(* IEC 61131-3 sources: CS_4_Aufzugsteuerung/src/Stations/CP112/Steuerung/Class/SdiasSafetyManagerFSoE (part 2) *)

            LastRequest := _WriteSysTime;

            //copy SDO into write-buffer
            ToStdLib.MemCpy(dest := #p_Handle_SDO_Write^.SDOStructure, source := #StandardRequest, size := (sizeof(SDOHeader.StdHeader.CRC) + StandardRequest.SDOHeader.Len));

            //mark SDO data as valid
            p_Handle_SDO_Write^.us_Status := SAFETY_SDO_DATA_VALID;

            if ( pISafety^.udVersion >= 16#1001 ) then
              SAFETY_iPushSafetyTask();
            end_if;

            SDOTimeMark       := ops.tAbsolute;
            ud_LastSetSysTime := ops.tAbsolute;
            eResponseState    := _wait;

            // check timeout
          elsif ((ops.tAbsolute - SDOTimeMark) > SDIAS_SAFTEY_SDO_RESPONSE_TIMEOUT) & (eResponseState <> _valid) then
            LogError("@029F (SdiasSafetyManagerFSoE::InitModule) Timeout while waiting for the SDO Send buffer to get ready (set system time)");
            eInitSSWErrorStep := eInitSSW;
            eInitSSW          := _InitError;
          end_if;

      //*****************************************************
        _wait: // wait for response

          //check id sdo sending was ok
          if ( p_Handle_SDO_Read^.us_Status = SAFETY_SDO_DATA_VALID ) then

            //calculate length of SDO
            us_SDO_length := sizeof(SDOHeader.StdHeader.CRC) + p_Handle_SDO_Read^.SDOStructure.SDOHeader.StdHeader.Len;

            //copy SDO without first byte (=status byte)
            ToStdLib.MemCpy(dest := p_SDOOutputBuffer, source := #p_Handle_SDO_Read^.SDOStructure, size := us_SDO_length );

            //mark data as received
            p_Handle_SDO_Read^.us_Status := SAFETY_SDO_NO_DATA;

            //check, if it's our answer
            if ((p_SDOOutputBuffer^.SDOHeader.StdHeader.Typ$USINT AND SBF_SSDO_MASK_TYPE)$t_SafetyFrameType = SDO_STD) then
              StandardResponse := (p_SDOOutputBuffer$^StandardFrameType)^;
              if StandardResponse.SDOHeader.SeqNr = (StandardSeqNr OR 16#80) then
                if LastRequest = _WriteSysTime then
                  // delete request
                  LastRequest           := _NoOpenRequest;
                  ud_AsyComRetryCounter := 0; // reset retry counter
                  eResponseState        := _valid;
                  // if returnvalue is 34 (E_SM_SSDO_INVALID_VIRTADDR) the virtual address is not supported by firmware
                  if StandardResponse.aData[0] <> 34 then
                    //virtual adress for write of timestamp is supported
                    b_SetSysTime := TRUE;
                  else
                    b_SetSysTime := FALSE;
                  end_if;
                else
                  LogError("@025A (SdiasSafetyManagerFSoE::InitModule) SDO Receive: Invalid standard frame response.");
                  eInitSSWErrorStep := eInitSSW;
                  eInitSSW          := _InitError;
                end_if;

                // if request is deleted, increase sequence number to set next request
                if LastRequest = _NoOpenRequest then
                  if StandardSeqNr < 16#7F then
                    StandardSeqNr += 1;
                  else
                    StandardSeqNr := 0;
                  end_if;
                end_if;
              else
                LogError("@025B (SdiasSafetyManagerFSoE::InitModule) SDO Receive: Invalid sequence number in Standard SDO response.");
                LogValue("expected: 0x{0} / received: 0x{1}", Value:=(StandardSeqNr OR 16#80), Value2:=StandardResponse.SDOHeader.SeqNr);
                eInitSSWErrorStep := eInitSSW;
                eInitSSW          := _InitError;
              end_if;
            else
              // ignore non-standard frames => the module may try to distribute it's configuration
            end_if;
          end_if;

          // check timeout
          if ((ops.tAbsolute - SDOTimeMark) > SDIAS_SAFTEY_SDO_RESPONSE_TIMEOUT) & (eResponseState <> _valid) then
            LogError("@02A1 (SdiasSafetyManagerFSoE::InitModule) SDO Response timeout while waiting for the module configuration.");
            eInitSSWErrorStep := eInitSSW;
            eInitSSW          := _InitError;
          end_if;
      //*****************************************************
        _valid:
          eInitSSW        := _DisablePLL;
          eResponseState  := _idle;
      //*****************************************************
      end_case;

//**********************************************************************************************************************************************************
    _DisablePLL: // disable the PLL
      TmpRetCode := BusConfigWrite(Offset:=SDIAS_SAFETY_PLL_OFFSET + t_PllRegister.StatusControl, Length:=sizeof(sPllRegister.StatusControl), pData:=#sPllRegister.StatusControl, IsControlAccess:=TRUE);

      if TmpRetCode = READY then
        eInitSSW := _GetPLLSettings;
      elsif TmpRetCode = ERROR then
        eInitSSW := _InitError;
      end_if;

//**********************************************************************************************************************************************************
    _GetPLLSettings: // get the actual PLL settings
      TmpRetCode := BusConfigRead(Offset:=SDIAS_SAFETY_PLL_OFFSET, Length:=sizeof(sPllRegister), pData:=#sPllRegister, IsControlAccess:=TRUE);

      if TmpRetCode = READY then
        // get bus cycle time for the PLL settings
        MyPara.uiCmd     := _BUS_IF_GET_BUSCYCLE_TIME;

        ToBusInterface.NewInst(pPara:=#MyPara, pResult:=#MyResult);
        if MyResult.aData[0]$t_GetBusCycleTime.retcode = _BUS_IF_RETVAL_OK then
          udBusTime       := MyResult.aData[0]$t_GetBusCycleTime.udBusCycleTime;
        else
          // use this just to have
          udBusTime := 1000;
          LogError("@02AA (SdiasSafetyManagerFSOE::InitModule) Failed to get bus cycle settings BusInterface.");
        end_if;

        udBusTime_us := udBusTime / 1000;

        // settings for pll
        sPllRegister.SystemPeriodTime           := udBusTime / 10;            // convert to 10*ns
        sPllRegister.StatusControl              := 0;
        sPllRegister.StatusControl.SyncEnable   := 1;
        sPllRegister.PeriodDivider              := to_usint(udBusTime_us / 1000);  // Bustime / 1ms to get divider (0 and 1 gets the same result)
        //sPllRegister.CompensationDelay // Keep value
        sPllRegister.SyncOut0.Offset            := 0;
        sPllRegister.SyncOut0.PeriodMultiplier  := to_usint(1000 / udBusTime_us);  // 1ms / Bustime to get multiplier (0 and 1 gets the same result);
        sPllRegister.SyncOut0.SyncStartDelay    := 0;
        sPllRegister.SyncOut0.ControlStatusRegister.SyncOutEnable     := 1;
        sPllRegister.SyncOut0.ControlStatusRegister.StartDelayEnable  := 0;
        if sPllRegister.PeriodDivider <= 1 then
          // no divider use system sync
          sPllRegister.SyncOut0.ControlStatusRegister.SyncSelector       := 1;  // no divider use system sync
        else
          // a divider is defined -> use it
          sPllRegister.SyncOut0.ControlStatusRegister.SyncSelector       := 0;
        end_if;

        eInitSSW := _ConfigurePLL;
      elsif TmpRetCode = ERROR then
        eInitSSW := _InitError;
      end_if;

//**********************************************************************************************************************************************************
    _ConfigurePLL:
      TmpRetCode := BusConfigWrite(Offset:=SDIAS_SAFETY_PLL_OFFSET, Length:=sizeof(sPllRegister), pData:=#sPllRegister, IsControlAccess:=TRUE);

      if TmpRetCode = READY then

        eInitSSW := _ConfigureTripleBufferAnalogReadData;
      elsif TmpRetCode = ERROR then
        eInitSSW := _InitError;
      end_if;

//**********************************************************************************************************************************************************
    _ConfigureTripleBufferAnalogReadData:

      //check if config from triple buffer for analog data is necessary
      if usAnalogInputByteSize then

        // configure the triple buffer - the required bytes are passed to the FPGA.
        sAnalogTripleBufferConfig.usSizeuCtoCPU := usAnalogInputByteSize - sizeof(USINT); //-1 byte for messagecounter
        sAnalogTripleBufferConfig.usSizeCPUtouC := 0; //Analog write when supported

        TmpRetCode := BusConfigWrite(Offset:=SBF_OFFSET_ANALOG_VALUE_TRIPLE_PUFFER_SWITCH_OFFSET_WR_1, Length:=sizeof(sAnalogTripleBufferConfig), pData:=#sAnalogTripleBufferConfig, IsControlAccess:=FALSE);

        if TmpRetCode = READY then
          eInitSSW := _ConfigureFastTripleBuffer;
        elsif TmpRetCode = ERROR then
          eInitSSW := _InitError;
        end_if;
      else
        eInitSSW := _ConfigureFastTripleBuffer;
      end_if;

//**********************************************************************************************************************************************************
    _ConfigureFastTripleBuffer:

      //check if init from triple buffer is necessary
      if uiPDOReadSizeFastUnsafeVar <> 0 |
        uiPDOWriteSizeFastUnsafeVar <> 0 then

        // configure the triple buffer - the required bytes are passed to the FPGA.
        sFastTripleBufferConfig.SizeuCtoCPU := uiPDOReadSizeFastUnsafeVar$USINT - 1;
        sFastTripleBufferConfig.SizeCPUtouC := uiPDOWriteSizeFastUnsafeVar$USINT - 1;

        TmpRetCode := BusConfigWrite(Offset:=SBF_OFFSET_FAST_UNSAFE_BUFFER_CONFIG, Length:=sizeof(sFastTripleBufferConfig), pData:=#sFastTripleBufferConfig, IsControlAccess:=FALSE);

        if TmpRetCode = READY then
          eInitSSW := _Finished;
        elsif TmpRetCode = ERROR then
          eInitSSW := _InitError;
        end_if;
      else
        eInitSSW := _Finished;
      end_if;

//**********************************************************************************************************************************************************
    _Finished:
      //Only set online here to 1 if we don't have to adjust the the triple buffer config, otherwise online will be set in cyclic after correcting the triple buffer config
      if b_ModuleAccessReady & (bWriteAnalogTripleBufferConfig = FALSE) then
        Online := 1;
      end_if;

      eInitSSW          := _PrepareInit;
      ModuleInitState   := READY;

#ifdef SAFETY_iDisableNonClassCommunication
      if ( pISafety^.udVersion >= 16#1002 ) then
        SAFETY_iDisableNonClassCommunication(uiMaster:=0, pucNode:=p_ObjectPath, uiDisable:=0);
      end_if;
#endif

//**********************************************************************************************************************************************************
    _InitError:
      eInitSSW          := _PrepareInit;
      ModuleInitState   := ERROR;

#ifdef SAFETY_iDisableNonClassCommunication
      if ( pISafety^.udVersion >= 16#1002 ) then
        SAFETY_iDisableNonClassCommunication(uiMaster:=0, pucNode:=p_ObjectPath, uiDisable:=0);
      end_if;
#endif

//**********************************************************************************************************************************************************
  end_case;

END_FUNCTION

FUNCTION VIRTUAL GLOBAL SdiasSafetyManagerFSoE::ClassSvr::NewInst
  VAR_INPUT
    pPara 	: ^CmdStruct;
    pResult 	: ^results;
  END_VAR
  VAR_OUTPUT
    ret_code 	: iprStates;
  END_VAR
  VAR
    i                 : UDINT;
    pSafetyModuleInfo : ^t_SdiasSafetyModuleInfo;
    MyPara 	          : CmdStruct;
    MyResult          : Results;
    HBGPlace          : UDINT;
    bRequiredError    : BOOL;
    bHWConfigError    : BOOL;

    pStr_HWTRequested     : ^CHAR;
    tmpplace      : USINT;
    pStr_HWTreeEntry : ^CHAR;
    usNextPlace   : USINT;
    pNewElement   : t_pHWCGetHardwareDiagnosisOutDynExt;
    usTmpAnalogInputByteSize : USINT;
  END_VAR

  ret_code := ERROR;

  CASE pPara^.uiCmd OF

//*****************************************************************************
//**  COMMANDS FROM BUS INTERFACE                                            **
//*****************************************************************************

//**********************************************************************************************************************************************************
    _BUS_IF_INIT_ACCESSES:
      // is called until the module is ready or in error state (only done once when no accesses have been created yet)
      ret_code := InitAccess();

//**********************************************************************************************************************************************************
    _BUS_IF_INIT_MODULE:
      // is called until the module is ready or in error state (done every time the module is connected)
      ret_code := InitModule();

//**********************************************************************************************************************************************************
    _BUS_IF_SDO_RESPONSE:
      // check if the command matches the one we're waiting for
      if (pPara^.aPara[0] = LastSDO.Command) &
         (pPara^.aPara[1] = LastSDO.Offset)  &
         (pPara^.aPara[2] = LastSDO.Length) then

        if pPara^.aPara[3]$iprStates = READY then
          if (LastSDO.Command = _BUS_IF_READ_VIA_SDO) then
            if (LastSDO.Offset = SBF_OFFSET_IO_MODULE_IDS) then
              if eResponseState = _wait then
                if pPara^.aPara[5] = LastSDO.Length then
                  if pPara^.aPara[4] then
                    // all parameters are fine, so we're ready
                    ret_code := READY;

                    _memcpy(ptr1:=#aModuleIDs, ptr2:=pPara^.aPara[4]$pVoid, cntr:=LastSDO.Length);

                    bRequiredError := FALSE;
                    bHWConfigError := FALSE;

                    //Set byte size of analog inputs to zero (will be summarized with every analog module)
                    usTmpAnalogInputByteSize := 0;

                    // search for a HBG in the module IDs
                    HBGPlace := SDIAS_SAFETY_INVALID_MAX_PLACE;
                    for i := 0 to 16 do
                      if (aModuleIDs[i] AND SDIAS_SAFETY_MODULE_ID_BUS_MASK) = SDIAS_SAFETY_MODULE_ID_CAN_BUS_MASK then
                        HBGPlace := i;
                        exit;
                      end_if;
                    end_for;

                    // now we got the module IDs according to the safety cpu => check if it matches our configuration (only available on newer firmware versions)
                    if b_GotOptionalSettings then
                      pSafetyModuleInfo := #aSafetyModuleInfo[0];

                      // always the same command
                      MyPara.uiCmd := SDIAS_SET_CLASS_STATE;

                      for i := 0 to 15 do
                        MyPara.aPara[1] := aModuleIDs[i];

                        // if a required module is not matching => required error
                        if pSafetyModuleInfo^.sdRequired & (aModuleIDs[i] <> pSafetyModuleInfo^.usExpectedDeviceID) then
                          MyPara.aPara[0] := _RequiredError$DINT;
                          bRequiredError := TRUE;
                          if aModuleIDs[i] = SDIAS_SAFETY_INVALID_DEVICE_ID then
                            LogValue("@02AB (SdiasSafetyManagerFSoE::ClassSvr::NewInst) No safety IO module at required place {0}", Value:=i);
                          else
                            LogValue("@02AC (SdiasSafetyManagerFSoE::ClassSvr::NewInst) Wrong safety IO module at required place {0}", Value:=i);
                          end_if;

                        // check if the configuration in the safety designer matches the configuration in the hardware classes
                        elsif pSafetyModuleInfo^.usExpectedDeviceID = OptionalSettings.ModuleIDsConfigured[i] then
                          // if it's an invalid device ID, it's only allowed if there is no module
                          if pSafetyModuleInfo^.usExpectedDeviceID = SDIAS_SAFETY_INVALID_DEVICE_ID then
                            if aModuleIDs[i] = SDIAS_SAFETY_INVALID_DEVICE_ID then
                              // correct (no module configured and no module found)
                              MyPara.aPara[0] := _ClassOk$DINT;  // this value is not being written to the module since if the ID is 0, there is also no this pointer to call the newinst
                            elsif (i <> HBGPlace) then
                              // no module configured but a module has been found at this place
                              LogValue("@02AD (SdiasSafetyManagerFSoE::ClassSvr::NewInst) No module configured in hardware classes and safety designer but found module at place {0}", Value:=i);
                              MyPara.aPara[0] := _WrongHardware$DINT; // again no object to write this value to
                              bHWConfigError := TRUE;
                            end_if;

                          // now check if we got the expected ID at this position
                          elsif aModuleIDs[i] = pSafetyModuleInfo^.usExpectedDeviceID then
                            // correct module
                            MyPara.aPara[0] := _ClassOk$DINT;

                            //Check if this is an analog module
                            if pSafetyModuleInfo^.usAnalogInputByteSize then
                              //Increase our byte size --> mabye we need to refresh the byte size in the tripple buffer of the analog values if the amount of configured modules
                              //differs to the amount of available modules on the hardware (e.g optional modules)
                              if usTmpAnalogInputByteSize = 0 then
                                usTmpAnalogInputByteSize += pSafetyModuleInfo^.usAnalogInputByteSize + sizeof(USINT);  //Add one byte for message counter if not added yet (first byte of analog input buffer is messagecounter)
                              else
                                usTmpAnalogInputByteSize += pSafetyModuleInfo^.usAnalogInputByteSize;
                              end_if;
                            end_if;

                            // if this module is optional
                          elsif OptionalSettings.OptionalFlagsIOModules AND (1 SHL i) then
                            // if it's a blank module
                            if aModuleIDs[i] = SDIAS_SAFETY_MODULE_ID_BLANK_MODULE then
                              // ok: blank is allowed at optional place
                              MyPara.aPara[0] := _NoHardware$DINT;

                              // don't send the blank-module ID
                              MyPara.aPara[1] := SDIAS_SAFETY_INVALID_DEVICE_ID;
                            else
                              if aModuleIDs[i] = SDIAS_SAFETY_INVALID_DEVICE_ID then
                                // ok: no module instead of the configured one (allowed since it's the last module. no more modules possible after an invalid device id)
                                MyPara.aPara[0] := _NoHardware$DINT;

                              //optional module, maybe this module is the HBG itself
                              elsif (HBGPlace <> SDIAS_SAFETY_INVALID_MAX_PLACE) & (i = HBGPlace) then

                                //OK: optional module is not available and this one is the HBG
                                MyPara.aPara[0] := _NoHardware$DINT;
                                MyPara.aPara[1] := SDIAS_SAFETY_INVALID_DEVICE_ID;
                              else
                                // wrong module detected
                                MyPara.aPara[0] := _WrongHardware$DINT;
                                bHWConfigError := TRUE;
                                LogValue("@02AE (SdiasSafetyManagerFSoE::ClassSvr::NewInst) Wrong safety IO module at place {0}. (configured as optional)", Value:=i);
                              end_if;
                            end_if;
                          else
                            // the module id does not match (missing or wrong module)
                            if aModuleIDs[i] = SDIAS_SAFETY_INVALID_DEVICE_ID then
                              MyPara.aPara[0] := _NoHardware$DINT;
                            else
                              MyPara.aPara[0] := _WrongHardware$DINT;
                            end_if;

                            // check if it's required
                            if MyPara.aPara[0] = _NoHardware$DINT then
                              LogValue("@02AF (SdiasSafetyManagerFSoE::ClassSvr::NewInst) No safety IO module at place {0}.", Value:=i);
                            else
                              LogValue("@02B0 (SdiasSafetyManagerFSoE::ClassSvr::NewInst) Wrong safety IO module at place {0}.", Value:=i);
                            end_if;

                            bHWConfigError := TRUE;
                          end_if;
                        else
                          // the configuration in the safety designer differs from the configuration via the hardware classes

                          // if the available hardware matches the safety designer configuration and there is no module (only in hw class configuration)
                          if (OptionalSettings.ModuleIDsConfigured[i] = SDIAS_SAFETY_INVALID_DEVICE_ID) &
                             ((aModuleIDs[i] = SDIAS_SAFETY_INVALID_DEVICE_ID) | (i = HBGPlace)) &
                             (pSafetyModuleInfo^.usExpectedDeviceID <> SDIAS_SAFETY_INVALID_DEVICE_ID) then
                            // that's allowed
                            LogValue("@02B1 (SdiasSafetyManagerFSoE::ClassSvr::NewInst) Module in hardware class configuration which is neither available physically nor in safety designer configuration at place {0}", Value:=i);
                            MyPara.aPara[0] := _NoHardware$DINT;

                          else
                            // in all other cases, it isn't
                            LogValue("@02B2 (SdiasSafetyManagerFSoE::ClassSvr::NewInst) Module in hardware class configuration differs from safety designer configuration at place {0}", Value:=i);
                            MyPara.aPara[0] := _InvalidConfguration$DINT;
                            bHWConfigError := TRUE;
                          end_if;
                        end_if;

                        if pSafetyModuleInfo^.pThis then
                          pSafetyModuleInfo^.pThis^.NewInst(#MyPara, #MyResult);
                        end_if;

                        pSafetyModuleInfo += sizeof(t_SdiasSafetyModuleInfo);
                      end_for;

                      //Check if our calculated size differs to the set one --> there must be optional analog modules which are not available
                      //So we need to set the size of the triple buffer config again, otherwise it won't work
                      if usTmpAnalogInputByteSize <> usAnalogInputByteSize then
                        usAnalogInputByteSize := usTmpAnalogInputByteSize;
                        bWriteAnalogTripleBufferConfig := TRUE;
                      end_if;

                      // check for hbg
                      if sHBG.pThis then
                        CanActive := OldCanActive := FALSE;
                        MyPara.uiCmd := SDIAS_SET_CLASS_STATE;

                        if HBGPlace <> SDIAS_SAFETY_INVALID_MAX_PLACE then
                          MyPara.aPara[1] := aModuleIDs[HBGPlace];

                          // if it's the wrong module and it's required => required error
                          if sHBG.sdRequired & (aModuleIDs[HBGPlace] <> sHBG.usExpectedDeviceID) then
                            MyPara.aPara[0] := _RequiredError$DINT;
                            bRequiredError := TRUE;
                            LogError("@02B3 (SdiasSafetyManagerFSoE::ClassSvr::NewInst) Wrong safety CAN terminal found instead of the configured required module!");

                          elsif (OptionalSettings.ModuleIDHBG = sHBG.usExpectedDeviceID) then
                            // the configured ID of LASAL and safety designer are equal

                            // if the module ID found is also the same => everthing is fine
                            if aModuleIDs[HBGPlace] = sHBG.usExpectedDeviceID then
                              MyPara.aPara[0] := _ClassOk$DINT;
                              CanActive := OldCanActive := TRUE;
                            else
                              // found something else
                              LogError("@02B4 (SdiasSafetyManagerFSoE::ClassSvr::NewInst) Wrong safety CAN terminal found (config of safety designer and hw classes match)");
                              MyPara.aPara[0] := _WrongHardware$DINT;
                              bHWConfigError := TRUE;
                            end_if;
                          else
                            // configuration of safety designer and hw classes does not match
                            LogError("@02B5 (SdiasSafetyManagerFSoE::ClassSvr::NewInst) Safety CAN terminal in hardware class configuration differs from safety designer configuration.");
                            MyPara.aPara[0] := _InvalidConfguration$DINT;
                            bHWConfigError := TRUE;
                          end_if;
                        else
                          MyPara.aPara[1] := SDIAS_SAFETY_INVALID_DEVICE_ID;

                          // projected in LASAL but not found in hardware
                          if sHBG.sdRequired then
                            MyPara.aPara[0] := _RequiredError$DINT;
                            bRequiredError := TRUE;
                            LogError("@02B6 (SdiasSafetyManagerFSoE::ClassSvr::NewInst) Required safety CAN terminal not available!");
                          else
                            // module is configured in safety designer
                            if (OptionalSettings.ModuleIDHBG <> SDIAS_SAFETY_INVALID_DEVICE_ID) then
                              // if the configuration does not match with the hardware classes
                              if (OptionalSettings.ModuleIDHBG <> sHBG.usExpectedDeviceID) then
                                LogError("@02B5 (SdiasSafetyManagerFSoE::ClassSvr::NewInst) Safety CAN terminal in hardware class configuration differs from safety designer configuration.");
                                MyPara.aPara[0] := _InvalidConfguration$DINT;
                                bHWConfigError := TRUE;

                              // the IDs match but it's not optional. since it's not available => error
                              elsif (OptionalSettings.OptionalFlagHBG.1 = FALSE) then
                                MyPara.aPara[0] := _NoHardware$DINT;
                                LogError("@02B7 (SdiasSafetyManagerFSoE::ClassSvr::NewInst) Could not find the non-optional Safety CAN terminal defined in the safety designer configuration.");
                                bHWConfigError := TRUE;

                              else
                                // if the IDs match and it's optional => just show no hardware (no error)
                                MyPara.aPara[0] := _NoHardware$DINT;
                              end_if;
                            else
                              LogError("@02B8 (SdiasSafetyManagerFSoE::ClassSvr::NewInst) Safety CAN terminal in hardware class configuration but not physically available and not in safety designer configuration.");
                              MyPara.aPara[0] := _NoHardware$DINT;
                            end_if;
                          end_if;
                        end_if;
                        sHBG.pThis^.NewInst(#MyPara, #MyResult);
                      else
                        // nothing projected for HBG in the lasal project

                        // if module is configured in safety designer
                        if (OptionalSettings.ModuleIDHBG <> SDIAS_SAFETY_INVALID_DEVICE_ID) then
                          // if a HBG has been found
                          if HBGPlace <> SDIAS_SAFETY_INVALID_MAX_PLACE then
                            // if it's not the configured module
                            if (aModuleIDs[HBGPlace] <> OptionalSettings.ModuleIDHBG) then
                              LogError("@02B9 (SdiasSafetyManagerFSoE::ClassSvr::NewInst) Safety CAN terminal found doesn't match the safety designer configuration.");
                              bHWConfigError := TRUE;
                            end_if;
                          else
                            // module not available (only a problem if it's not optional)
                            if (OptionalSettings.OptionalFlagHBG.1 = FALSE) then
                              LogError("@02BA (SdiasSafetyManagerFSoE::ClassSvr::NewInst) Could not find the non-optional Safety CAN terminal defined in the safety designer configuration.");
                              bHWConfigError := TRUE;
                            end_if;
                          end_if;
                        else
                          // module not configured in safety designer. if there is a module available, the number of IOs in safety does not match the config
                          if HBGPlace <> SDIAS_SAFETY_INVALID_MAX_PLACE then
                            LogError("@02BB (SdiasSafetyManagerFSoE::ClassSvr::NewInst) Safety CAN terminal found but not projected in the safety designer configuration.");
                            bHWConfigError := TRUE;
                          end_if;
                        end_if;
                      end_if;
                    else
                      // old firmware (no optional settings available)
                      if MaxPlace <> SDIAS_SAFETY_INVALID_MAX_PLACE then
                        pSafetyModuleInfo := #aSafetyModuleInfo[0];

                        // always the same command
                        MyPara.uiCmd := SDIAS_SET_CLASS_STATE;

                        for i := 0 to MaxPlace do
                          if pSafetyModuleInfo^.pThis then
                            MyPara.aPara[1] := aModuleIDs[i];
                            if aModuleIDs[i] = pSafetyModuleInfo^.usExpectedDeviceID then
                              MyPara.aPara[0] := _ClassOk$DINT;
                            elsif aModuleIDs[i] <> SDIAS_SAFETY_INVALID_DEVICE_ID then
                              if pSafetyModuleInfo^.sdRequired then
                                MyPara.aPara[0] := _RequiredError$DINT;
                                bRequiredError := TRUE;
                                LogValue("@02AC (SdiasSafetyManagerFSoE::ClassSvr::NewInst) Wrong safety IO module at required place {0}.", Value:=i);
                              else
                                MyPara.aPara[0] := _WrongHardware$DINT;
                                bHWConfigError  := TRUE;
                              end_if;
                            else
                              if pSafetyModuleInfo^.sdRequired then
                                MyPara.aPara[0] := _RequiredError$DINT;
                                bRequiredError := TRUE;
                                LogValue("@02AB (SdiasSafetyManagerFSoE::ClassSvr::NewInst) No safety IO module at required place {0}.", Value:=i);
                              else
                                MyPara.aPara[0] := _NoHardware$DINT;
                                // Hardwareclass placed in Project but no physical Hardware available is allowed
                                // bHWConfigError  := TRUE;
                              end_if;
                            end_if;
                            pSafetyModuleInfo^.pThis^.NewInst(#MyPara, #MyResult);

                          elsif aModuleIDs[i] <> SDIAS_SAFETY_INVALID_DEVICE_ID then  // HWK this pointer is NIL but a module is identified
                            bHWConfigError  := TRUE;
                          end_if;

                          pSafetyModuleInfo += sizeof(t_SdiasSafetyModuleInfo);
                        end_for;
                      end_if;

                      // Check if a module info was passed for which there is no corrosponding HWK object.
                      if MaxPlace + 1 < sizeof(t_ModuleIDs) then
                        // it's only a config error if it's not the HBG
                        if (aModuleIDs[MaxPlace + 1] <> SDIAS_SAFETY_INVALID_DEVICE_ID) & ((MaxPlace + 1) <> HBGPlace) then
                          bHWConfigError  := TRUE;
                        end_if;
                      end_if;

                      // check for hbg
                      if sHBG.pThis then
                        MyPara.uiCmd := SDIAS_SET_CLASS_STATE;
                        if HBGPlace <> SDIAS_SAFETY_INVALID_MAX_PLACE then
                          MyPara.aPara[1] := aModuleIDs[HBGPlace];

                          if aModuleIDs[HBGPlace] = sHBG.usExpectedDeviceID then
                            MyPara.aPara[0] := _ClassOk$DINT;
                            CanActive := OldCanActive := TRUE;
                            bHWConfigError := FALSE;
                          elsif aModuleIDs[HBGPlace] <> SDIAS_SAFETY_INVALID_DEVICE_ID then
                            if sHBG.sdRequired then
                              MyPara.aPara[0] := _RequiredError$DINT;
                              bRequiredError := TRUE;
                              LogError("@02BE (SdiasSafetyManagerFSoE::ClassSvr::NewInst) Wrong safety IO module at required HBG place.");
                            else
                              MyPara.aPara[0] := _WrongHardware$DINT;
                              CanActive := OldCanActive := FALSE;
                            end_if;
                          else
                            if sHBG.sdRequired then
                              MyPara.aPara[0] := _RequiredError$DINT;
                              bRequiredError := TRUE;
                              LogError("@02BF (SdiasSafetyManagerFSoE::ClassSvr::NewInst) HBG required but not available!");
                            else
                              MyPara.aPara[0] := _NoHardware$DINT;
                              CanActive := OldCanActive := FALSE;
                            end_if;
                          end_if;
                        else
                          MyPara.aPara[1] := SDIAS_SAFETY_INVALID_DEVICE_ID;
                          if sHBG.sdRequired then
                            MyPara.aPara[0] := _RequiredError$DINT;
                            bRequiredError := TRUE;
                            LogError("@02BE (SdiasSafetyManagerFSoE::ClassSvr::NewInst) Wrong safety IO module at required HBG place.");
                          else
                            MyPara.aPara[0] := _WrongHardware$DINT;
                            CanActive := OldCanActive := FALSE;
                          end_if;
                        end_if;
                        sHBG.pThis^.NewInst(#MyPara, #MyResult);
                      end_if;
                    end_if;

                    if bRequiredError then
                      MyPara.uiCmd := _BUS_IF_SET_REQUIRED_ERROR;
                      ToBusInterface.NewInst(#MyPara, #MyResult);
                    end_if;

                    if bHWConfigError then
                      // if we have optional settings, we already logged the reason
                      if b_GotOptionalSettings = FALSE then
                        LogError("@02C0 (SdiasSafetyManagerFSoE::ClassSvr::NewInst) Hardwareconfiguration does not match objects placed in network.");
                      end_if;

                      // Check if Safetymanyger is required
                      MyPara.uiCmd     := _BUS_IF_GET_REQUIRED_SETTING;
                      ToBusInterface.NewInst(pPara:=#MyPara, pResult:=#MyResult);
                      if MyResult.aData[0]$t_BusIFRetvalErrorcode = _BUS_IF_RETVAL_OK then
                        // if it's required => set required error
                        if MyResult.aData[4] then

                          MyPara.uiCmd := _BUS_IF_SET_REQUIRED_ERROR;
                          ToBusInterface.NewInst(#MyPara, #MyResult);
                        else

                          SetSafetyState(_WrongSafetyHW);
                          Online      := 0;

                          // Update BusIF ClassState
                          MyPara.uiCmd := _BUS_IF_SET_CLASS_STATE;
                          MyPara.aPara[0] := _WrongHardware$DINT;
                          ToBusInterface.NewInst(#MyPara, #MyResult);

                          // Cancel init
                          eInitSSWErrorStep := eInitSSW;
                          eInitSSW := _InitError;

                          // Set Module states
                          pSafetyModuleInfo := #aSafetyModuleInfo[0];
                          // always the same command
                          MyPara.uiCmd := SDIAS_SET_CLASS_STATE;
                          MyPara.aPara[0] := _ModuleFoundButManagerIsOff$DINT;

                          if MaxPlace <> SDIAS_SAFETY_INVALID_MAX_PLACE then
                            for i := 0 to MaxPlace do
                              if pSafetyModuleInfo^.pThis then
                                MyPara.aPara[1] := aModuleIDs[i];
                                pSafetyModuleInfo^.pThis^.NewInst(#MyPara, #MyResult);
                              end_if;
                              pSafetyModuleInfo += sizeof(t_SdiasSafetyModuleInfo);
                            end_for;
                          end_if;

                          // check for hbg
                          if sHBG.pThis then
                            sHBG.pThis^.NewInst(#MyPara, #MyResult);
                          end_if;

                        end_if;

                      end_if;

                    end_if;

                  else
                    LogError("@02C1 (SdiasSafetyManagerFSoE::ClassSvr::NewInst) Invalid SDO response buffer pointer.");
                  end_if;
                else
                  LogError("@02C2 (SdiasSafetyManagerFSoE::ClassSvr::NewInst) Invalid length for SDO response data.");
                end_if;

                eResponseState := _valid;
              else
                LogError("@02C3 (SdiasSafetyManagerFSoE::ClassSvr::NewInst) SDO response arrived when no response was expected.");
              end_if;
            end_if;
          elsif (LastSDO.Command = _BUS_IF_WRITE_VIA_SDO) then

              ret_code := READY;

              // we got the response to our write memory access
              LastSDO.ResponseArrived := TRUE;

          elsif (LastSDO.Command = _BUS_IF_READ_VIA_SDO_CTRL) then
            if LastSDO.ResponseArrived = FALSE then
              if pPara^.aPara[5] = LastSDO.Length then
                if pPara^.aPara[4] then
                  // all parameters are fine, so we're ready
                  ret_code := READY;

                  // copy the response data
                  _memcpy(ptr1:=Config.pActData, ptr2:=pPara^.aPara[4]$pVoid, cntr:=LastSDO.Length);
                else
                  LogError("@02C1 (SdiasSafetyManagerFSoE::ClassState::NewInst) Invalid SDO response buffer pointer.");
                end_if;
              else
                LogError("@02C2 (SdiasSafetyManagerFSoE::ClassState::NewInst) Invalid length for SDO response data.");
              end_if;

              LastSDO.ResponseArrived := TRUE;
            else
              LogError("@02C3 (SdiasSafetyManagerFSoE::ClassState::NewInst) SDO response arrived when no response was expected.");
            end_if;
          elsif (LastSDO.Command = _BUS_IF_WRITE_VIA_SDO_CTRL) then
            if LastSDO.ResponseArrived = FALSE then
              // all parameters are fine, so we're ready
              ret_code := READY;

              LastSDO.ResponseArrived := TRUE;
            else
              LogError("@02C3 (SdiasSafetyManagerFSoE::ClassState::NewInst) SDO response arrived when no response was expected.");
            end_if;
          end_if;
        else
          LogError("@02C4 (SdiasSafetyManagerFSoE::ClassSvr::NewInst) SDO transfer failed.");
        end_if;
      else
        LogError("@02C5 (SdiasSafetyManagerFSoE::ClassSvr::NewInst) Received invalid SDO response.");
      end_if;

//**********************************************************************************************************************************************************
    _BUS_IF_DATA_POINTER_AVAILABLE:
      // does nothing in the FSoE version
      ret_code := READY;

//**********************************************************************************************************************************************************
    _BUS_IF_RESET_DETECTED:
      // don't overwrite other errors
      if SafetyState = _SafetyClassOK then
        SafetyState := _LostPowerSupply;
      end_if;

      // check if module is requred
      MyPara.uiCmd     := _BUS_IF_GET_REQUIRED_SETTING;
      ToBusInterface.NewInst(pPara:=#MyPara, pResult:=#MyResult);
      if MyResult.aData[0]$t_BusIFRetvalErrorcode = _BUS_IF_RETVAL_OK then
        // if it's required => set required error
        if MyResult.aData[4] then

          MyPara.uiCmd := _BUS_IF_SET_REQUIRED_ERROR;
          ToBusInterface.NewInst(#MyPara, #MyResult);
        end_if;
      end_if;

      // drop config of connected modules

      // initialize the message for the periphery
      MyPara.uiCmd := SDIAS_SET_CLASS_STATE;
      MyPara.aPara[1] := 0;// no device ID
      MyPara.aPara[0] := _NoHardware$DINT;

      // tell the connected IO module objects
      if MaxPlace <> SDIAS_SAFETY_INVALID_MAX_PLACE then
        pSafetyModuleInfo := #aSafetyModuleInfo[0];

        for i := 0 to MaxPlace do
          if pSafetyModuleInfo^.pThis then
            pSafetyModuleInfo^.pThis^.NewInst(#MyPara, #MyResult);
          end_if;

          pSafetyModuleInfo += sizeof(t_SdiasSafetyModuleInfo);
        end_for;
      end_if;

      // tell the hbg (if available)
      if sHBG.pThis then
        sHBG.pThis^.NewInst(#MyPara, #MyResult);
      end_if;

//**********************************************************************************************************************************************************
    _BUS_IF_RESET_GONE_DETECTED:
      if SafetyState = _LostPowerSupply then

        // get safety and serial numbers of connected modules
        bUpdateModuleConfig := TRUE;

        // remember the time. in case we don't get the SDO response to signal the firmware being ready, we use a timeout
        ud_ResetGoneTime := ops.tAbsolute;

        // we wait for an asynchronous SDO response in the cyclic of the base class. once we got that, the firmware is ready
        b_WaitForFirmwareBoot := TRUE;

        // refetch IDs of connected modules
        eCheckIDSSW := _Wait4Idle;

        SafetyState := _SafetyClassOK;
      end_if;

//**********************************************************************************************************************************************************

    CMD_GET_HARDWARE_DIAGNOSIS:
      //Returns module info
      ret_code := ERROR;
      pResult^.aData[0]$t_HWCGetHardwareDiagnosisOut.retcode := _HWC_RETVAL_ERROR;

      pStr_HWTRequested := pPara^.aPara[0]$t_HWCGetHardwareDiagnosisIn.pStr_HardewareTreeEntry;

      tmpplace := (pStr_HWTRequested+pPara^.aPara[0]$t_HWCGetHardwareDiagnosisIn.us_current_index)^$USINT;

      //Check if pointer is valid
      if aSafetyModuleInfo[tmpplace].pThis then

        // Set Offline Device ID
        pResult^.aData[0]$t_HWCGetHardwareDiagnosisOut.ud_DeviceID := (aSafetyModuleInfo[tmpplace].usExpectedDeviceID AND 2#00111000 ) shr 3;   // Bit 3-5 Modul typ
        pResult^.aData[0]$t_HWCGetHardwareDiagnosisOut.ud_Variante :=  aSafetyModuleInfo[tmpplace].usExpectedDeviceID AND 2#00000111;  // Bit 0-2 Submodul typ

        if aModuleIDs[tmpplace] = aSafetyModuleInfo[tmpplace].usExpectedDeviceID then

          ret_code := READY;
          pResult^.aData$t_HWCGetHardwareDiagnosisOut.retcode := _HWC_RETVAL_OK;

          pResult^.aData[0]$t_HWCGetHardwareDiagnosisOut.ud_DeviceID  := (aModuleIDs[tmpplace] AND 2#00111000 ) shr 3;  // Bit 3-5 Modul typ
          pResult^.aData[0]$t_HWCGetHardwareDiagnosisOut.ud_Variante  :=  aModuleIDs[tmpplace] AND 2#00000111; // // Bit 0-2 Submodul typ
          pResult^.aData[0]$t_HWCGetHardwareDiagnosisOut.ud_Place     := tmpplace;
          pResult^.aData[0]$t_HWCGetHardwareDiagnosisOut.hd_HWVersion :=  sHwVersions.aVersion[tmpplace];  //Hardware version of module

          //Get firmware version of module (if available)
          GetFWVersion(udPlace:=tmpplace, pData:=#a_FWVersion[0],sizeof(a_FWVersion));
          pResult^.aData$t_HWCGetHardwareDiagnosisOut.pStr_FWVersion := #a_FWVersion[0];

          // Get Serialno ---------------------------------------------------------------------------------------------
          _memcpy(ptr1 := #a_SerialNo[0]
                , ptr2 := #sSafetySerNrs.aSerialNumbers[tmpplace]
                , cntr := sizeof(sSafetySerNrs.aSerialNumbers[tmpplace]) );

          a_SerialNo[sizeof(sSafetySerNrs.aSerialNumbers[tmpplace])] := 0;  // 0 Terminierung

          pResult^.aData[0]$t_HWCGetHardwareDiagnosisOut.pStr_SerialNo := #a_SerialNo[0];

          pResult^.aData[0]$t_HWCGetHardwareDiagnosisOut.hd_SafetyNumber  := sSafetySerNrs.aSafetyNumbers[tmpplace];

          // first free the old then create the memory (linked list) for the additional information

          if pAdditionalDiagInfo then
            HwDiagFreeDynExtList(pList:=pAdditionalDiagInfo);
          end_if;
          pAdditionalDiagInfo      := NIL;

          // add the firmware version
          pNewElement := HwDiagAddDynExt2List(ppList:=#pAdditionalDiagInfo, EntryID:=_HWC_DIAG_ID_SAFETY_FIRMWARE_VERSION, udVersion:=1, udDataLength:=sizeof(HDINT));

          if pNewElement then
            // add the data in the reserved memory
            (pNewElement$^HDINT + sizeof(t_HWCGetHardwareDiagnosisOutDynExt))^ := FirmwareVersion;
          end_if;

          // add the safety designer project name
          pNewElement := HwDiagAddDynExt2List(ppList:=#pAdditionalDiagInfo, EntryID:=_HWC_DIAG_ID_SAFETY_DESIGNER_PROJECT_NAME, udVersion:=1, udDataLength:=ProjectNameStr.GetLength());

          if pNewElement then
            // add the data in the reserved memory
            ProjectNameStr.ReadDataOff(udOff:=0, pData:=pNewElement$^USINT + sizeof(t_HWCGetHardwareDiagnosisOutDynExt), udMax:=pNewElement^.ud_DataLength);
          end_if;

          // add the safety designer project revision
          pNewElement := HwDiagAddDynExt2List(ppList:=#pAdditionalDiagInfo, EntryID:=_HWC_DIAG_ID_SAFETY_DESIGNER_PROJECT_REVISION, udVersion:=1, udDataLength:=ProjectRevisionStr.GetLength());

          if pNewElement then
            // add the data in the reserved memory
            ProjectRevisionStr.ReadDataOff(udOff:=0, pData:=pNewElement$^USINT + sizeof(t_HWCGetHardwareDiagnosisOutDynExt), udMax:=pNewElement^.ud_DataLength);
          end_if;

          pResult^.aData[0]$t_HWCGetHardwareDiagnosisOut.p_DynExtList := pAdditionalDiagInfo;

        elsif aModuleIDs[tmpplace] <> SDIAS_SAFETY_INVALID_DEVICE_ID then
          pResult^.aData$t_HWCGetHardwareDiagnosisOut.retcode := _HWC_RETVAL_ERROR_WRONG_HARDWARE;
        else
          pResult^.aData$t_HWCGetHardwareDiagnosisOut.retcode := _HWC_RETVAL_ERROR_NO_HARDWARE;
        end_if;

      else
        pResult^.aData[0]$t_HWCGetHardwareDiagnosisOut.retcode := _HWC_RETVAL_ERROR_SDIAS_MODULE_NOT_FOUND;
      end_if;

//**********************************************************************************************************************************************************
    CMD_GET_HARDWARE_TREE_ENTRY:
      //Returns module info

      ret_code := ERROR;
      pResult^.aData[0]$t_HWCGetHardwareTreeEntryOut.retcode := _HWC_RETVAL_ERROR;

      pStr_HWTreeEntry := pPara^.aPara[0]$t_HWCGetHardwareTreeEntryIn.pStr_LastHardewareTreeEntry;

      //First HWT Path
      if (pStr_HWTreeEntry + pStr_HWTreeEntry$^UINT^)^ <> HWT_ESCAPE_INTERNALBUS_SDIAS_SAFETY then  // + 1 for Byte length -1 for 2nd last element of string

        if aSafetyModuleInfo[0].pThis then

          _memcpy(ptr1 := #a_HWTEntryStr[0]
                , ptr2 := pPara^.aPara[0]$t_HWCGetHardwareTreeEntryIn.pStr_LastHardewareTreeEntry
                , cntr := pPara^.aPara[0]$t_HWCGetHardwareTreeEntryIn.pStr_LastHardewareTreeEntry$^UINT^ +2 );  // +2 2 Byte Strlength is not included in the stringlength

          // Add escape sequence
          a_HWTEntryStr[0]$UINT += 1;
          a_HWTEntryStr[a_HWTEntryStr[0]$UINT+1] := HWT_ESCAPE_INTERNALBUS_SDIAS_SAFETY;

          // Add Place
          a_HWTEntryStr[0]$UINT += 1;
          a_HWTEntryStr[a_HWTEntryStr[0]$UINT+1] := 0;

          //Return Hardware Tree Entry and set return codes
          pResult^.aData[0]$t_HWCGetHardwareTreeEntryOut.pStr_NextHardewareTreeEntry := #a_HWTEntryStr[0];

          pResult^.aData[0]$t_HWCGetHardwareTreeEntryOut.retcode := _HWC_RETVAL_OK_HWTSTR_RETURNED;
          ret_code := READY;

        else
          pResult^.aData[0]$t_HWCGetHardwareTreeEntryOut.retcode := _HWC_RETVAL_ERROR_SDIAS_MODULE_NOT_FOUND;
        end_if;

      //search next module
      else

        usNextPlace := (pStr_HWTreeEntry  + pPara^.aPara[0]$t_HWCGetHardwareTreeEntryIn.us_current_index)^$USINT+1;

        if usNextPlace <= SDIAS_SAFETY_MAX_PLACE_NR &
           aSafetyModuleInfo[usNextPlace].pThis then

          _memcpy(ptr1 := #a_HWTEntryStr[0]
                , ptr2 := pPara^.aPara[0]$t_HWCGetHardwareTreeEntryIn.pStr_LastHardewareTreeEntry
                , cntr := pPara^.aPara[0]$t_HWCGetHardwareTreeEntryIn.pStr_LastHardewareTreeEntry$^UINT^ +2 );  // +2 2 Byte Strlength is not included in the stringlength

          // Set new Place
          a_HWTEntryStr[a_HWTEntryStr[0]$UINT + 1] := usNextPlace;

          pResult^.aData[0]$t_HWCGetHardwareTreeEntryOut.pStr_NextHardewareTreeEntry := #a_HWTEntryStr[0];

          //Return Hardware Tree Entry and set return codes
          pResult^.aData[0]$t_HWCGetHardwareTreeEntryOut.retcode := _HWC_RETVAL_OK_HWTSTR_RETURNED;
          ret_code := READY;

        else
          ret_code := READY;
          pResult^.aData$t_HWCGetHardwareTreeEntryOut.retcode := _HWC_RETVAL_OK_END_OF_LIST;
        end_if;
      end_if;

//**********************************************************************************************************************************************************

//*****************************************************************************
//** INTERNAL COMMANDS                                                       **
//*****************************************************************************

//**********************************************************************************************************************************************************
    CMD_SM_READ_PDO_SIZE:
      // get the size of the PDO
      LastSDO.Command := _BUS_IF_READ_VIA_SDO;
      LastSDO.Offset  := SBF_OFFSET_SPDO_LENGTH;
      LastSDO.Length  := sizeof(UINT);

      MyPara.uiCmd    := LastSDO.Command$UINT;
      MyPara.aPara[0] := LastSDO.Offset;
      MyPara.aPara[1] := LastSDO.Length;
      ret_code := ToBusInterface.NewInst(#MyPara, #MyResult);

//**********************************************************************************************************************************************************
  else
    ret_code := SafetyBaseFSoE::NewInst(pPara, pResult);
//**********************************************************************************************************************************************************
  END_CASE;

END_FUNCTION

FUNCTION VIRTUAL SdiasSafetyManagerFSoE::ShowProjectRevision

  ProjectNameStr.WriteDataOff(udLen:=PrjNameStrLen + 1, udOff:=0, pData:=pPrjNameStr);

  ProjectRevisionStr.WriteDataOff(udLen:=PrjRevStrLen + 1, udOff:=0, pData:=pPrjRevStr);

END_FUNCTION

FUNCTION VIRTUAL SdiasSafetyManagerFSoE::InitSafeModule
  VAR_OUTPUT
    sd_retval 	: DINT;
  END_VAR

  // allocate memory for finding unsafe-IO-Servers
  // in first place we allocate 512 byte for our blocked transfers
  p_BlockedTransferMemory := ToStdLib.Malloc( size := SBF_CONFIG_MEMORY_BLOCK_SIZE );
  IF p_BlockedTransferMemory <> NIL THEN
    ud_BlockedTransferMemorySize := SBF_CONFIG_MEMORY_BLOCK_SIZE;
  ELSE
    SafetyState := _MemAllocFailed;
    sd_retval := -100;
    return;
  END_IF;

  // if there is a safety manager to gather the configuration
  if pSafetyManagerThis then
    // allocate memory for gathering configuration information => in first place we allocate 512 byte
    pConfigMem := ToStdLib.Malloc( size := SBF_CONFIG_MEMORY_BLOCK_SIZE );
    IF pConfigMem <> NIL THEN
      ConfigMemSize := SBF_CONFIG_MEMORY_BLOCK_SIZE;
      ConfigMemSizeUsed := 4;
    ELSE
      SafetyState := _MemAllocFailed;
      sd_retval := -100;
      return;
    END_IF;
  end_if;

END_FUNCTION

FUNCTION VIRTUAL GLOBAL SdiasSafetyManagerFSoE::CanOut::NewInst
  VAR_INPUT
    pPara 	: ^CmdStruct;
    pResult 	: ^results;
  END_VAR
  VAR_OUTPUT
    ret_code 	: iprStates;
  END_VAR
  VAR
    tempCmd         : CmdStruct;
    _result         : results;
  END_VAR

  ret_code := ERROR;  //Default is error

  CASE pPara^.uiCmd OF
//**********************************************************************************************************************************************************
    SDIAS_SAFETY_LOGIN_HBG:
      // check parameters
      if pPara^.aPara[0] & pPara^.aPara[1] then

        ret_code := READY;  //Parameters are ok, set retcode

        sHBG.pThis               := pPara^.aPara[0]$pVirtualBase;
        sHBG.usExpectedDeviceID  := pPara^.aPara[1]$USINT;
        sHBG.sdRequired          := pPara^.aPara[2];
        sHBG.pIOStates           := pPara^.aPara[3]$^HDINT;

        // if leds/hgb not added so far, add them
        if StateBytesUsed = 0 then
          StateBitsUsed := (sizeof(t_LedAndIOStates.biLEDs) + sizeof(t_LedAndIOStates.HBGInputs)) * 8;
          // refresh state bytes used value
          StateBytesUsed := ((StateBitsUsed-1) / 8) + 1;
        end_if;

        if sHBG.sdRequired & (b_AnyModuleRequired = FALSE) then
          b_AnyModuleRequired := TRUE;
          // if any access is required => the businterface is also required
          tempCmd.uiCmd := _BUS_IF_SET_REQUIRED;
          ToBusInterface.NewInst(pPara:=#tempCmd, pResult:=#_result);
          if _result.aData[0]$t_BusIFRetvalErrorcode <> _BUS_IF_RETVAL_OK then
            LogError("@029D (SdiasSafetyManagerFSoE::CanOut::NewInst) Failed to set the BusInterface to required.");
          end_if;
        end_if;
      end_if;
//**********************************************************************************************************************************************************
  END_CASE;

END_FUNCTION

FUNCTION VIRTUAL SdiasSafetyManagerFSoE::GetConfiguration
  VAR
    pHelp                 : ^void;
    SizeToGo              : UINT;
    ActSize               : UINT;
    ActAddr               : HDINT;
    SDOReqBuf             : SDORequReadConfig;
    SDORspBuf             : ARRAY [0..SBF_SDO_MAX_LENGTH-1] OF USINT;
    pRspBuf               : ^SDORespReadConfig;
    i                     : DINT;
    pSafetyModuleInfo     : ^t_SdiasSafetyModuleInfo;
    MyPara 	              : CmdStruct;
    MyResult              : Results;
  END_VAR

  //initialize header-data for request

  //calculate length without crc
  SDOReqBuf.StdHeader.Len := sizeof(SDORequReadConfig) - sizeof(SDOHeader.StdHeader.CRC);

  //type
  SDOReqBuf.StdHeader.Typ := SDO_STD;

  //command for reading config data
  SDOReqBuf.StdHeader.Cmd := SBF_SDO_COMMAND_READ;

  // read the complete 256 Bytes of safety and serial number info
  pHelp    := #sSafetySerNrs;
  SizeToGo := sizeof(sSafetySerNrs);
  pRspBuf  := (#SDORspBuf)$^SDORespReadConfig;
  ActAddr  := SBF_SDO_ADDRESS_SER_NR_DATA;

  while SizeToGo do
    if SizeToGo > SDIAS_SAFTEY_SDO_MAX_DATA_PER_PAKET then
      ActSize := SDIAS_SAFTEY_SDO_MAX_DATA_PER_PAKET;
    else
      ActSize := SizeToGo;
    end_if;

    if SDOReadCfgRequ(p_SDORequestBuffer  := #SDOReqBuf,
                      p_SDOResponseBuffer := pRspBuf,
                      ud_Address          := ActAddr,
                      us_Length           := ActSize$USINT,
                      b_UseCache          := FALSE) then
      LogError("@02C6 (SdiasSafetyManagerFSoE::GetConfiguration) Failed to get safety and serial numbers of the IO modules.");
      return;
    else
      _memcpy(ptr1:=pHelp, ptr2:=#pRspBuf^.ud_Data, cntr:=ActSize);
    end_if;

    SizeToGo  -= ActSize;
    ActAddr   += ActSize;
    pHelp     += ActSize;
  end_while;

  // read the complete 64 Bytes of hardware version info
  pHelp    := #sHwVersions;
  SizeToGo := sizeof(sHwVersions);
  pRspBuf  := (#SDORspBuf)$^SDORespReadConfig;
  ActAddr  := SBF_SDO_ADDRESS_HW_VERSIONS;

  while SizeToGo do
    if SizeToGo > SDIAS_SAFTEY_SDO_MAX_DATA_PER_PAKET then
      ActSize := SDIAS_SAFTEY_SDO_MAX_DATA_PER_PAKET;
    else
      ActSize := SizeToGo;
    end_if;

    if SDOReadCfgRequ(p_SDORequestBuffer  := #SDOReqBuf,
                      p_SDOResponseBuffer := pRspBuf,
                      ud_Address          := ActAddr,
                      us_Length           := ActSize$USINT,
                      b_UseCache          := FALSE) then
      LogError("@02F9 (SdiasSafetyManagerFSoE::GetConfiguration) Failed to get hw versions of the Safe IO modules!");
      return;
    else
      // if the return code in the response buffer is not 0 => the virtual memory is not available
      if pRspBuf^.us_Returncode <> 0 then
        // reset array to make sure there are no hw versions stored
        _memset(dest:=#sHwVersions.aVersion[0], usByte:=0, cntr:=sizeof(sHwVersions));
        exit;
      end_if;

      _memcpy(ptr1:=pHelp, ptr2:=#pRspBuf^.ud_Data, cntr:=ActSize);
    end_if;

    SizeToGo  -= ActSize;
    ActAddr   += ActSize;
    pHelp     += ActSize;
  end_while;

  // check if the firmware version info is availble
  if sFirmwareVersion.RevMinor >= SBF_FW_VER_FW_INFO_AVAILABLE then

    // read the complete 64 Bytes of firmware version info
    pHelp    := #sFWVersions;
    SizeToGo := sizeof(sFWVersions);
    pRspBuf  := (#SDORspBuf)$^SDORespReadConfig;
    ActAddr  := SBF_SDO_ADDRESS_HW_VERSIONS + sizeof(sHwVersions); //After the hw version, there is a 64 byte block with the fw version of each module

    while SizeToGo do
      if SizeToGo > SDIAS_SAFTEY_SDO_MAX_DATA_PER_PAKET then
        ActSize := SDIAS_SAFTEY_SDO_MAX_DATA_PER_PAKET;
      else
        ActSize := SizeToGo;
      end_if;

      if SDOReadCfgRequ(p_SDORequestBuffer  := #SDOReqBuf,
                        p_SDOResponseBuffer := pRspBuf,
                        ud_Address          := ActAddr,
                        us_Length           := ActSize$USINT,
                        b_UseCache          := FALSE) then
        LogError("@0790 (SdiasSafetyManagerFSoE::GetConfiguration) Failed to get fw versions of the Safe IO modules!");
        return;
      else
        // if the return code in the response buffer is not 0 => the virtual memory is not available
        if pRspBuf^.us_Returncode <> 0 then
          // reset array to make sure there are no fw versions stored
          _memset(dest:=#sFWVersions.aVersion[0], usByte:=0, cntr:=sizeof(sFWVersions));
          exit;
        end_if;

        _memcpy(ptr1:=pHelp, ptr2:=#pRspBuf^.ud_Data, cntr:=ActSize);
      end_if;

      SizeToGo  -= ActSize;
      ActAddr   += ActSize;
      pHelp     += ActSize;
    end_while;

  end_if;

  // only available for IOs, not the HBG
  if MaxPlace <> SDIAS_SAFETY_INVALID_MAX_PLACE then
    // always the same command
    MyPara.uiCmd := SDIAS_SET_NUMBERS;

    pSafetyModuleInfo := #aSafetyModuleInfo[0];
    for i := 0 to MaxPlace$DINT do
      // safety number
      MyPara.aPara[0] := (sSafetySerNrs.aSafetyNumbers[i])$DINT;

      // pointer to serial number string
      MyPara.aPara[1] := (#sSafetySerNrs.aSerialNumbers[i][0])$DINT;

      // hw version
      MyPara.aPara[2] := (sHwVersions.aVersion[i])$DINT;

      // fw version
      MyPara.aPara[3] := (sFWVersions.aVersion[i])$DINT;

      if pSafetyModuleInfo^.pThis then
        pSafetyModuleInfo^.pThis^.NewInst(#MyPara, #MyResult);
      end_if;

      pSafetyModuleInfo += sizeof(t_SdiasSafetyModuleInfo);
    end_for;
  end_if;

END_FUNCTION

FUNCTION VIRTUAL GLOBAL SdiasSafetyManagerFSoE::DisconnectEvent
  VAR
    i                 : UDINT;
    pSafetyModuleInfo : ^t_SdiasSafetyModuleInfo;
    MyPara 	          : CmdStruct;
    MyResult          : Results;
  END_VAR

  SafetyBaseFSoE::DisconnectEvent();

  // initialize the message for the periphery
  MyPara.uiCmd := SDIAS_SET_CLASS_STATE;
  MyPara.aPara[1] := 0;// no device ID
  MyPara.aPara[0] := _NoHardware$DINT;

  // tell the connected IO module objects
  if MaxPlace <> SDIAS_SAFETY_INVALID_MAX_PLACE then
    pSafetyModuleInfo := #aSafetyModuleInfo[0];

    for i := 0 to MaxPlace do
      if pSafetyModuleInfo^.pThis then
        pSafetyModuleInfo^.pThis^.NewInst(#MyPara, #MyResult);
      end_if;

      pSafetyModuleInfo += sizeof(t_SdiasSafetyModuleInfo);
    end_for;
  end_if;

  // tell the hbg (if available)
  if sHBG.pThis then
    sHBG.pThis^.NewInst(#MyPara, #MyResult);
  end_if;

  // clear the strings
  ProjectNameStr.Clear();
  ProjectRevisionStr.Clear();

END_FUNCTION

FUNCTION VIRTUAL SdiasSafetyManagerFSoE::SetSafetyState
  VAR_INPUT
    NewState 	: SafetyConfigStateType;
  END_VAR
  VAR
    MyPara 	  : CmdStruct;
    MyResult	: results;
  END_VAR

  // use it locally
  SafetyState := NewState;

  // tell the outer class
  MyPara.uiCmd := SDIAS_SET_SAFETY_STATE;
  MyPara.aPara[0] := NewState$DINT;
  ToBusInterface.NewInst(#MyPara, #MyResult);

END_FUNCTION

FUNCTION VIRTUAL GLOBAL SdiasSafetyManagerFSoE::CyWork
  VAR_INPUT
    EAX 	: UDINT;
  END_VAR
  VAR_OUTPUT
    state (EAX) 	: UDINT;
  END_VAR
  VAR
    MyPara 	          : CmdStruct;
    MyResult          : Results;
    TmpRetCode        : iprStates;
  END_VAR

  if bWriteAnalogTripleBufferConfig then

    // configure the triple buffer - the required bytes are passed to the FPGA.
    if usAnalogInputByteSize = 0 then
      sAnalogTripleBufferConfig.usSizeuCtoCPU := 0; //no analog data used
    else
      sAnalogTripleBufferConfig.usSizeuCtoCPU := usAnalogInputByteSize - sizeof(USINT); //-1 byte for messagecounter
    end_if;

    sAnalogTripleBufferConfig.usSizeCPUtouC := 0; //Analog write when supported

    TmpRetCode := BusConfigWrite(Offset:=SBF_OFFSET_ANALOG_VALUE_TRIPLE_PUFFER_SWITCH_OFFSET_WR_1, Length:=sizeof(sAnalogTripleBufferConfig), pData:=#sAnalogTripleBufferConfig, IsControlAccess:=FALSE);

    if TmpRetCode = READY then
      bWriteAnalogTripleBufferConfig := FALSE;
      if b_ModuleAccessReady then
        //Set online, because we now have set the correct offset for the triple buffer to switch
        Online := 1;
      end_if;

    elsif TmpRetCode = ERROR then
      bWriteAnalogTripleBufferConfig := FALSE;
      LogError("@08A4 (SdiasSafetyManagerFSoE::CyWork) Failed to configure triple buffer for analog input data.");
    end_if;
  end_if;

  // if the initialisiation has been finished and there is an object for the hbg check if it's has been connected or disconnected
  if Online then

    case eCheckIDSSW of
  //**********************************************************************************************************************************************************
      _Nothing:
        if sHBG.pThis then
          // check for a can connect event
          if CanActive > OldCanActive then
            // if we're already idle => get it on
            if eResponseState = _idle then
              eCheckIDSSW := _GetIDs;
            else
              // otherwise, wait for it (need to remember the connect event)
              eCheckIDSSW := _Wait4Idle;
            end_if;

          // check for a can disconnect event
          elsif CanActive < OldCanActive then
            if sHBG.sdRequired then
              // if it's required => required error
              MyPara.uiCmd := _BUS_IF_SET_REQUIRED_ERROR;
              ToBusInterface.NewInst(#MyPara, #MyResult);
            else
              // otherwise show that it has been disconnected
              MyPara.uiCmd := SDIAS_SET_CLASS_STATE;
              MyPara.aPara[1] := 0;// no device ID
              MyPara.aPara[0] := _NoHardware$DINT;
              sHBG.pThis^.NewInst(#MyPara, #MyResult);
            end_if;
          end_if;
          OldCanActive := CanActive;
        end_if;

  //**********************************************************************************************************************************************************
      _Wait4Idle:
        if eResponseState = _idle then
          eCheckIDSSW := _GetIDs;
        end_if;

  //**********************************************************************************************************************************************************
      _GetIDs:
        case eResponseState of
        //*****************************************************
          _idle:
            LastSDO.Command := _BUS_IF_READ_VIA_SDO;
            LastSDO.Offset  := SBF_OFFSET_IO_MODULE_IDS;
            LastSDO.Length  := sizeof(t_ModuleIDs);

            MyPara.uiCmd    := LastSDO.Command$UINT;
            MyPara.aPara[0] := LastSDO.Offset;
            MyPara.aPara[1] := LastSDO.Length;
            TmpRetcode := ToBusInterface.NewInst(#MyPara, #MyResult);
            if TmpRetcode = READY then
              SDOTimeMark  := ops.tAbsolute;
              eResponseState:= _wait;
            elsif TmpRetcode = ERROR then
              LogError("@02A7 (SdiasSafetyManagerFSoE::InitModule) Failed to add read SDO for module configuration.");
            end_if;
        //*****************************************************
          _wait:
            // wait for response
            if ((ops.tAbsolute - SDOTimeMark) > SDIAS_SAFTEY_SDO_RESPONSE_TIMEOUT) then
              LogError("@02A1 (SdiasSafetyManagerFSoE::InitModule) SDO Response timeout while waiting for the module configuration.");
              eCheckIDSSW := _Nothing;
              eResponseState := _idle;
            end_if;
        //*****************************************************
          _valid:
            eCheckIDSSW := _Nothing;
            eResponseState := _idle;
        //*****************************************************
        end_case;
  //**********************************************************************************************************************************************************
    end_case;
  end_if;

  state := SafetyBaseFSoE::CyWork(0);

END_FUNCTION

FUNCTION VIRTUAL SdiasSafetyManagerFSoE::RefreshAsySrv
  VAR
    i                 : UDINT;
    pSafetyModuleInfo : ^t_SdiasSafetyModuleInfo;
    MyPara 	          : CmdStruct;
    MyResult          : Results;
    AsyValues         : t_AsyRefresh;
  END_VAR

  // tell the outer class
  MyPara.uiCmd := SDIAS_SET_ASY_STATE;
  AsyValues.QuitComError := QuitComError;
  MyPara.aPara[0] := (#AsyValues)$DINT;
  ToBusInterface.NewInst(#MyPara, #MyResult);

  // tell the connected IO module objects
  if MaxPlace <> SDIAS_SAFETY_INVALID_MAX_PLACE then
    pSafetyModuleInfo := #aSafetyModuleInfo[0];

    for i := 0 to MaxPlace do
      if pSafetyModuleInfo^.pThis then
        pSafetyModuleInfo^.pThis^.NewInst(#MyPara, #MyResult);
      end_if;

      pSafetyModuleInfo += sizeof(t_SdiasSafetyModuleInfo);
    end_for;
  end_if;

END_FUNCTION

FUNCTION VIRTUAL GLOBAL SdiasSafetyManagerFSoE::FastUnsafeOutputs::Write
  VAR_INPUT
    input (EAX) 	: BDINT;
  END_VAR
  VAR_OUTPUT
    result (EAX) 	: BDINT;
  END_VAR
  VAR
    pUnsafeOutLogin : ^t_FastUnsafeOuts;
  END_VAR

  // if the pointer is valid and we're in the first init run (the firstscan check prevents a crash caused by someone writing on the server during runtime)
  if input & (us_FirstScan < 2) then
    pUnsafeOutLogin := input$^t_FastUnsafeOuts;
    // check if it's the correct usage of the class
    if pUnsafeOutLogin^.Kennung = SDIAS_SAFETY_FAST_UNSAFE_KENNUNG then
      pFastUnsafeOutThis := pUnsafeOutLogin^.pThis;
    end_if;
  end_if;

  result := input;

END_FUNCTION

FUNCTION VIRTUAL GLOBAL SdiasSafetyManagerFSoE::FastUnsafeInputs::Write
  VAR_INPUT
    input (EAX) 	: BDINT;
  END_VAR
  VAR_OUTPUT
    result (EAX) 	: BDINT;
  END_VAR

  FastUnsafeInputs := input;
  result := FastUnsafeInputs;

END_FUNCTION

FUNCTION VIRTUAL SdiasSafetyManagerFSoE::SetRetryCounter
  VAR
    pSafetyModuleInfo : ^t_SdiasSafetyModuleInfo;
    MyPara 	 : CmdStruct;
    MyResult : Results;
    i        :  USINT;
  END_VAR

  if b_RetryCounterAvailable then

    if MaxPlace <> SDIAS_SAFETY_INVALID_MAX_PLACE then
      //Command for new inst call in sdiassafetybase
      MyPara.uiCmd := SDIAS_SET_RETRY_COUNTER;

      //calls newinst method of all safety modules which exists.
      for i := 0 to MaxPlace do
        pSafetyModuleInfo := #aSafetyModuleInfo[i];
        MyPara.aPara[0] := a_RetryCnt[i];
        MyPara.aPara[1] := a_RetryCnt[i+16];  //+16 for retry counter of µC2
        pSafetyModuleInfo^.pThis^.NewInst(#MyPara, #MyResult);
      end_for;
    end_if;
  else
    //Retrycounter not available -> show -1 at servers.
    SafetyRetryCounter := -1; //Not available

    if MaxPlace <> SDIAS_SAFETY_INVALID_MAX_PLACE then
      MyPara.uiCmd := SDIAS_RETRY_COUNTER_NOT_AVAILABLE;
      for i := 0 to MaxPlace do
        pSafetyModuleInfo := #aSafetyModuleInfo[i];
        pSafetyModuleInfo^.pThis^.NewInst(#MyPara, #MyResult);
      end_for;
    end_if;
  end_if;

END_FUNCTION

FUNCTION VIRTUAL GLOBAL SdiasSafetyManagerFSoE::Background
  VAR_INPUT
    EAX 	: UDINT;
  END_VAR
  VAR_OUTPUT
    state (EAX) 	: UDINT;
  END_VAR

  // if we have to update the module config, are not busy and the firmware has already booted (or a timeout on the boot occured)
  if bUpdateModuleConfig & (eCheckIDSSW = _Nothing) & ((b_WaitForFirmwareBoot = FALSE) | ((ops.tAbsolute - ud_ResetGoneTime) > SBF_FIRMWARE_BOOTUP_TIMEOUT)) then
    bUpdateModuleConfig := FALSE;

    GetConfiguration();
  end_if;

  state := SafetyBaseFSoE::Background(0);

END_FUNCTION

FUNCTION VIRTUAL SdiasSafetyManagerFSoE::BusConfigWrite
	VAR_INPUT
		Offset 	: HDINT;
		Length 	: UINT;
		pData 	: pVoid;
		IsControlAccess 	: BOOL;(* := FALSE *)
	END_VAR
	VAR_OUTPUT
		retcode 	: iprStates;
	END_VAR
  VAR
    TmpRetcode  : iprStates;
    MyPara      : CmdStruct;
    MyResult    : results;
  END_VAR

  retcode := BUSY;

  case Config.BusConfigSSW of
//**********************************************************************************************************************************************************
    _PrepareAccess:
      Config.RestLength := Length;
      Config.pActData   := pData;

      Config.BusConfigSSW := _StartAccess;

//**********************************************************************************************************************************************************
    _StartAccess:
      if IsControlAccess then
        LastSDO.Command := _BUS_IF_WRITE_VIA_SDO_CTRL;
      else
        LastSDO.Command := _BUS_IF_WRITE_VIA_SDO;
      end_if;

      LastSDO.Offset  := Offset$DINT;
      if Config.RestLength > SDIAS_SAFETY_MAX_SDO_DATA_PER_CYCLE then
        LastSDO.Length  := SDIAS_SAFETY_MAX_SDO_DATA_PER_CYCLE;
      else
        LastSDO.Length  := Config.RestLength;
      end_if;
      LastSDO.ResponseArrived := FALSE;

      MyPara.uiCmd    := LastSDO.Command;
      MyPara.aPara[0] := LastSDO.Offset;
      MyPara.aPara[1] := LastSDO.Length;
      MyPara.aPara[2] := Config.pActData$DINT;
      TmpRetcode := ToBusInterface.NewInst(#MyPara, #MyResult);
      if TmpRetcode = READY then
        Config.SDOTimeMark  := ops.tAbsolute;
        Config.BusConfigSSW := _Wait4Answer;
      elsif TmpRetcode = ERROR then
        retcode := ERROR;
        LogError("@02BC (SdiasSafetyManagerFSoE::BusConfigWrite) Failed to add write SDO for module configuration.");
      end_if;

//**********************************************************************************************************************************************************
    _Wait4Answer:
      // wait for response

      // check for response
      if LastSDO.ResponseArrived then
        Config.RestLength -= LastSDO.Length;
        Config.pActData   += LastSDO.Length;

        if Config.RestLength = 0 then
          retcode := READY;
          Config.BusConfigSSW := _PrepareAccess;
        end_if;
      elsif ((ops.tAbsolute - Config.SDOTimeMark) > SDIAS_SAFTEY_SDO_RESPONSE_TIMEOUT) then
        LogError("@02BD (SdiasSafetyManagerFSoE::BusConfigWrite) SDO Response timeout while waiting for the write response.");
        retcode := ERROR;
      end_if;

//**********************************************************************************************************************************************************
  end_case;

END_FUNCTION

FUNCTION VIRTUAL SdiasSafetyManagerFSoE::BusConfigRead
	VAR_INPUT
		Offset 	: HDINT;
		Length 	: UINT;
		pData 	: pVoid;
		IsControlAccess 	: BOOL;(* := FALSE *)
	END_VAR
	VAR_OUTPUT
		retcode 	: iprStates;
	END_VAR
  VAR
    TmpRetcode  : iprStates;
    MyPara      : CmdStruct;
    MyResult    : results;
  END_VAR

  retcode := BUSY;

  case Config.BusConfigSSW of
//**********************************************************************************************************************************************************
    _PrepareAccess:
      Config.RestLength := Length;
      Config.pActData   := pData;

      Config.BusConfigSSW := _StartAccess;

//**********************************************************************************************************************************************************
    _StartAccess:
      if IsControlAccess then
        LastSDO.Command := _BUS_IF_READ_VIA_SDO_CTRL;
      else
        LastSDO.Command := _BUS_IF_READ_VIA_SDO;
      end_if;

      LastSDO.Offset  := Offset$DINT;
      if Config.RestLength > SDIAS_SAFETY_MAX_SDO_DATA_PER_CYCLE then
        LastSDO.Length  := SDIAS_SAFETY_MAX_SDO_DATA_PER_CYCLE;
      else
        LastSDO.Length  := Config.RestLength;
      end_if;
      LastSDO.ResponseArrived := FALSE;

      MyPara.uiCmd    := LastSDO.Command;
      MyPara.aPara[0] := LastSDO.Offset;
      MyPara.aPara[1] := LastSDO.Length;
      TmpRetcode := ToBusInterface.NewInst(#MyPara, #MyResult);
      if TmpRetcode = READY then
        Config.SDOTimeMark  := ops.tAbsolute;
        Config.BusConfigSSW := _Wait4Answer;
      elsif TmpRetcode = ERROR then
        retcode := ERROR;
        LogError("@02BC (SdiasSafetyManagerFSoE::BusConfigRead) Failed to add write SDO for module configuration.");
      end_if;

//**********************************************************************************************************************************************************
    _Wait4Answer:
      // wait for response

      // check for response
      if LastSDO.ResponseArrived then
        Config.RestLength -= LastSDO.Length;
        Config.pActData   += LastSDO.Length;

        if Config.RestLength = 0 then
          retcode := READY;
          Config.BusConfigSSW := _PrepareAccess;
        end_if;
      elsif ((ops.tAbsolute - Config.SDOTimeMark) > SDIAS_SAFTEY_SDO_RESPONSE_TIMEOUT) then
        LogError("@02BD (SdiasSafetyManagerFSoE::BusConfigRead) SDO Response timeout while waiting for the write response.");
        retcode := ERROR;
      end_if;

//**********************************************************************************************************************************************************
  end_case;

END_FUNCTION

FUNCTION VIRTUAL SdiasSafetyManagerFSoE::HwDiagFreeDynExtList
	VAR_INPUT
		pList 	: ^t_HWCGetHardwareDiagnosisOutDynExt;
	END_VAR
  VAR
    pHelp 	: ^t_HWCGetHardwareDiagnosisOutDynExt;
  END_VAR

  while pList do
    // remember the current entry
    pHelp := pList;

    // set plist to the next entry and free pHelp
    pList := pList^.p_Next;

    // free the current entry
    ToStdLib.Free(mptr:=pHelp);
  end_while;

END_FUNCTION

FUNCTION VIRTUAL SdiasSafetyManagerFSoE::HwDiagAddDynExt2List
	VAR_INPUT
		ppList 	: ^t_pHWCGetHardwareDiagnosisOutDynExt;
		EntryID 	: t_HWCGetHardwareDiagnosisOutType;
		udVersion 	: UDINT;
		udDataLength 	: UDINT;
	END_VAR
	VAR_OUTPUT
		pNewElement 	: t_pHWCGetHardwareDiagnosisOutDynExt;
	END_VAR

  if ppList^ = NIL then
    ppList^$pVoid := ToStdLib.Malloc(size:=sizeof(t_HWCGetHardwareDiagnosisOutDynExt) + udDataLength);
    pNewElement := ppList^;
  else
    pNewElement := ppList^;
    while pNewElement^.p_Next <> NIL do
      pNewElement := pNewElement^.p_Next;
    end_while;
    pNewElement^.p_Next$pVoid := ToStdLib.Malloc(size:=sizeof(t_HWCGetHardwareDiagnosisOutDynExt) + udDataLength);
    pNewElement := pNewElement^.p_Next;
  end_if;

  if pNewElement <> NIL then
    // initialize the new memory
    pNewElement^.DiagID         := EntryID;
    pNewElement^.ud_Version     := udVersion;
    pNewElement^.p_Next         := NIL;
    pNewElement^.ud_DataLength  := udDataLength;

    if udDataLength then
      _memset(dest:=pNewElement + sizeof(t_HWCGetHardwareDiagnosisOutDynExt), usByte:=0, cntr:=udDataLength);
    end_if;
  end_if;

END_FUNCTION

FUNCTION VIRTUAL GLOBAL SdiasSafetyManagerFSoE::HGWOut::NewInst
  VAR_INPUT
    pPara 	: ^CmdStruct;
    pResult 	: ^Results;
  END_VAR
  VAR_OUTPUT
    ret_code 	: iprStates;
  END_VAR
  VAR
    tempCmd         : CmdStruct;
    _result         : results;
    dRetCode        : DINT;
  END_VAR

  ret_code := READY;

  case pPara^.uiCmd of

    //**********************************************************************************************************************************************************
    SDIAS_SAFETY_GET_HGW_INFO:

      //Check for valid version
      //*****************************************************************************
      if (pPara^.aPara[0] = 0x1) | (pPara^.aPara[0] = 0x2) then

        //Return version number
        pResult^.aData[0] := pPara^.aPara[0]$USINT;

        //pointer to input data to scp
        sHGW.pInputPDO           := pPara^.aPara[1]$^void;

        if sHGW.pInputPDO = nil then
          ret_code := ERROR;
          LogError(e_msg:="@03DD (SdiasSafetyManagerFSoE::HGWOut::NewInst) Pointer to input data of SCP is invalid.");
          return;
        end_if;

        // add PDO input data
        dRetCode := AddPDOToInputBuffer(ud_p2Buffer         := sHGW.pInputPDO$UDINT
                                      , ud_SafetyNr         := sHGW.hdSafetyNrb$UDINT
                                      , b_IsOptional        := FALSE
                                      , ui_PdoLen           := sHGW.InputPDOLength
                                      , ui_TargetOffset     := sHGW.InputPDOOffset
                                      );

        if dRetCode = -2 then
          //busy
          ret_code := BUSY;
          return;
        elsif dRetCode <> 0 then
          ret_code := ERROR;
          LogError(e_msg:="@072B (SdiasSafetyManagerFSoE::HGWOut::NewInst) Failed to add HGW PDO to input buffer.");
          return;
        end_if;

        // return the pointer to the Buffer (is linear local memory, so the offset can be added later)
        sHGW.pOutputPDO$UDINT := GetPointer2PDOBuffer();

        // here we have a difference depending on the version
        if pPara^.aPara[0] = 0x1 then

          pResult^.uiLng := 27;
          pResult^.aData[1]$UDINT := (sHGW.pOutputPDO+sHGW.OutputPDOOffset)$UDINT;
          pResult^.aData[5]$UINT  := sHGW.InputPDOLength;  //data to scp
          pResult^.aData[7]$UINT  := sHGW.OutputPDOLength; //data to hgw
          pResult^.aData[9]$UINT  := sHGW.uiSlotID;
          pResult^.aData[11]$UINT  := sHGW.uiCommunicationID;
          pResult^.aData[13]$USINT := sHGW.udMachineNrb$USINT;    //Old version, 1 byte machine number
          pResult^.aData[17]$USINT := sCPUConfig.CompPathLen$USINT;
          pResult^.aData[18]$UDINT := sCPUConfig.pCompPath$UDINT;
          pResult^.aData[22]$UDINT := sCPUConfig.SafetyNbr$UDINT;
          pResult^.aData[26]$UDINT := (#ErrorState)$UDINT;

        elsif pPara^.aPara[0] = 0x2 then

          pResult^.uiLng := 30;
          pResult^.aData[1]$UDINT := (sHGW.pOutputPDO+sHGW.OutputPDOOffset)$UDINT;
          pResult^.aData[5]$UINT  := sHGW.InputPDOLength;  //data to scp
          pResult^.aData[7]$UINT  := sHGW.OutputPDOLength; //data to hgw
          pResult^.aData[9]$UINT  := sHGW.uiSlotID;
          pResult^.aData[11]$UINT  := sHGW.uiCommunicationID;
          pResult^.aData[13]$UDINT := sHGW.udMachineNrb;
          pResult^.aData[17]$USINT := sCPUConfig.CompPathLen$USINT;
          pResult^.aData[18]$UDINT := sCPUConfig.pCompPath$UDINT;
          pResult^.aData[22]$UDINT := sCPUConfig.SafetyNbr$UDINT;
          pResult^.aData[26]$UDINT := (#ErrorState)$UDINT;

        end_if;

      //*****************************************************************************
      else
        // unknown version of the request
        ret_code := ERROR;
      end_if;

    //**********************************************************************************************************************************************************
    SDIAS_SAFETY_LOGIN_HGW:

      //Check for valid version
      if pPara^.aPara[0] = 0x1 then

      // check parameters
        if pPara^.aPara[1] then
          sHGW.pThis         := pPara^.aPara[1]$pVirtualBase; //this pointer of connect hgw communication class
          sHGW.sdRequired    := pPara^.aPara[2];              //required

        if sHGW.sdRequired & (b_AnyModuleRequired = FALSE) then
          b_AnyModuleRequired := TRUE;
          // if any access is required => the businterface is also required
          tempCmd.uiCmd := _BUS_IF_SET_REQUIRED;
          ToBusInterface.NewInst(pPara:=#tempCmd, pResult:=#_result);
          if _result.aData[0]$t_BusIFRetvalErrorcode <> _BUS_IF_RETVAL_OK then
            LogError("@03DE (SdiasSafetyManagerFSoE::HGWOut::NewInst) Failed to set the BusInterface to required");
          end_if;
        end_if;
      else
          ret_code := ERROR;
        end_if;

      else
        // unknown version of the request
        ret_code := ERROR;
      end_if;

    //**********************************************************************************************************************************************************
    CMD_SM_ADD_ROUTING_INFO:

      if sHGW.hdSafetyNrb <> pPara^.aPara[0]$HDINT then
        //safe act hgw safety number
        sHGW.hdSafetyNrb := pPara^.aPara[0]$HDINT;
        //add routing element for hgw panel
        dRetCode := AddRoutingElement(ud_SafeNumber:=sHGW.hdSafetyNrb, ud_thisp:=sHGW.pThis$UDINT, pPathInfo:=NIL);
        if dRetCode <> 0 then
          ret_code := ERROR;
        end_if;
      end_if;

    //**********************************************************************************************************************************************************
    CMD_SM_ADD_SDO_TO_BUFFER:
      ret_code := ClassSvr.NewInst(pPara:=pPara, pResult:=pResult);

  //**********************************************************************************************************************************************************

  else
    //if command is not known send it to safety manager
    if pSafetyManagerThis then
      ret_code := pSafetyManagerThis^.NewInst(pPara, pResult);
    end_if;

  end_case;

END_FUNCTION

FUNCTION VIRTUAL SdiasSafetyManagerFSoE::SafeActModuleConfig
  VAR_INPUT
    sActModuleConfig 	: t_ModuleCfg;
  END_VAR
  VAR
  	pCompPath : pVoid;
  END_VAR

  //only copy required information for HGW connection, see SDIAS_SAFETY_GET_HGW_INFO
  //do not copy pointers of paths, they point to a temporary memory. copy the content
  sCPUConfig.SafetyNbr := sActModuleConfig.SafetyNbr;
  if sCPUConfig.pCompPath then
    pCompPath := ToStdLib.ReAlloc(sCPUConfig.pCompPath, sActModuleConfig.CompPathLen);
  else
    pCompPath := ToStdLib.Malloc(sActModuleConfig.CompPathLen);
  end_if;
  if pCompPath then
    _memcpy(pCompPath, sActModuleConfig.pCompPath, sActModuleConfig.CompPathLen);
    sCPUConfig.pCompPath := pCompPath$^USINT;
    sCPUConfig.CompPathLen := sActModuleConfig.CompPathLen;
  end_if;

END_FUNCTION

FUNCTION VIRTUAL GLOBAL SdiasSafetyManagerFSoE::FCN_Command::Write
  VAR_INPUT
    input (EAX) 	: UDINT;
  END_VAR
  VAR_OUTPUT
    result (EAX) 	: UDINT;
  END_VAR

  // only if input is valid and we're in the right state
  if (input = 1) & (FCN_StateMachine = 1) then
    sFlexCon.CommandRequest := input;
  end_if;

  result := input;

END_FUNCTION

FUNCTION VIRTUAL SdiasSafetyManagerFSoE::GetFWVersion
	VAR_INPUT
    udPlace : UDINT;
		pData 	: ^CHAR;
		Length 	: UDINT;
	END_VAR

  //Returns the fw version of the Sdias IO modules behind the SCP

  //Check pointer
  if pData then
    //Length of Firmwareversion (HDINT) -> 8Byte +1 byte zero termination
    if Length >= 9 then
      //Check if fw version is available
      if sFWVersions.aVersion[udPlace] then
        _itoa(udNumber:=sFWVersions.aVersion[udPlace], pString:=pData);
      else
        pData^ := 0;  //No firmware version available
      end_if;
    else
      pData^ := 0;  //Invalid length
    end_if;
  end_if;

END_FUNCTION
